FUNCTION_BLOCK FB_Auslauf
VAR_INPUT
END_VAR
VAR_OUTPUT
END_VAR
VAR
END_VAR

IF GVL_IO.xLichtschranke_Auslauf AND GVL_IO.xServo_Auslauf_GS THEN
    GVL_IO.xAuslaufBereit := TRUE;
ELSIF NOT GVL_IO.xLichtschranke_Auslauf THEN
    GVL_IO.xAuslaufBereit := FALSE;
END_IF

END_FUNCTION_BLOCK

(* stored: Version 1.1.0.1
   POU FB_Auslauf: Id {a1863f5a-1c9a-45c2-b074-f03ce1135c66}, SpecialFunc None *)
